TYPE "ST_S11GraphProbe"
VERSION : 0.1
   STRUCT
      Go : Bool;
      Fault : Bool;
   END_STRUCT;
END_TYPE
